// TIA Portal V21 export
// export: Created 2026-11-10T07:35:04.8725218Z, ExportSetting WithDefaults, DisplayName Totally Integrated Automation Portal, DisplayVersion V21 Update 3, DisplayName STEP 7 Professional, DisplayVersion V21 Update 3, DisplayName STEP 7 Safety, DisplayVersion V21, DisplayName Tech WebApplication, DisplayVersion V21, DisplayName WinCC Basic/Comfort/Advanced, DisplayVersion V21 Update 3, DisplayName WinCC Unified, DisplayVersion V21 Update 3
FUNCTION_BLOCK "FB_Lad_ex043"   // FB18, LAD
{ S7_Optimized_Access := 'TRUE' }
VERSION : 0.1
// stored: AutoNumber true, IsIECCheckEnabled false, IsRetainMemResEnabled false, MemoryReserve 100, SetENOAutomatically false, UDAEnableTagReadback false
   VAR_INPUT
      v_part : PIP;
      v_ret_val : Int;
   END_VAR
   VAR_OUTPUT
      v_fladdr : Word;
   END_VAR
BEGIN

REGION Network 1: SYNC_PI - Synchronize the process image inputs
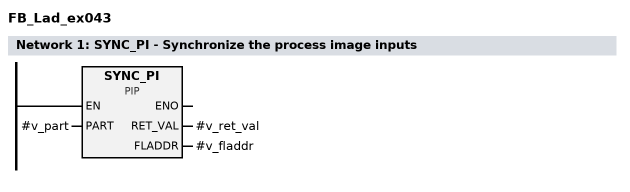
   RUNG wire#powerrail
      { S7_Templates := "value_type := PIP" } SYNC_PI(PART := #v_part, RET_VAL => #v_ret_val, FLADDR => #v_fladdr)
   END_RUNG
   // the same network as SCL:
   #v_ret_val := SYNC_PI(PART := #v_part, FLADDR => #v_fladdr);
END_REGION
END_FUNCTION_BLOCK
